Fanuc KAREL source: kt00016.KL

-- PROVISIONAL review KL for V940-1; original PC SHA256 82499ecc08bc44d66dd542690ba4f3cb5e484608f831ebc15742158b3d70d3b9
-- Incomplete behavior may be omitted. Consult companion uncertainty JSON. Do not deploy.
PROGRAM KT00016
%NOLOCKGROUP
VAR
  R1 : REAL
  OUT : REAL
-- UNRESOLVED_DECL H2 type=002017
BEGIN
  -- V9_ZERO_TABLE_METADATA_HINT layout=0001; no indexed target words; source/name/runtime held
  -- UNRESOLVED_PC offsets 5-16; opcodes 2E,23
  -- UNRESOLVED_PC offsets 21-35; opcodes 2E,22,9D,33,B4
  -- UNRESOLVED_PC offsets 40-63; opcodes 21,22,9D,33,B3,64,69,23
  -- UNRESOLVED_PC offsets 68-72; opcodes 7F
END KT00016
